{attribute 'qualified_only'}
{attribute 'strict'}
TYPE E_ResetHW :
(
	INIT := 0,
	RESET_HW := 10,
	DONE := 50
);
END_TYPE

(* stored: Version 1.1.0.1, ProductVersion 3.1.4024.12
   DUT E_ResetHW: Id {0d88b8cc-5541-4d33-9867-087aa81adb93} *)
